TYPE "ST_Nameplate"
VERSION : 0.1
   STRUCT
      ProductUri : WString[255];
      ManufacturerName : String[80];
      ProductDesignation : String[80];
      SerialNumber : String[40];
      YearOfConstruction : String[8];
      HardwareVersion : String[24];
      FirmwareVersion : String[24];
      SoftwareVersion : String[24];
      OrderCode : String[40];
      DocumentationUrl : WString[255];
   END_STRUCT;

END_TYPE

